Staubli VAL3: Force4Item.dtx

mdesc mNomSpeed
public string sArmType
public num nMaxJnt4Force[4]
